(* IEC 61131-3 sources: plc-st-coding-agent/progress/v13_r8/upstream/datasets/public/tests, 2 files *)

(* ---- public-easy-04.reference.st ---- *)
(* Numeric millisecond variant of the jam-pump task. DebounceMs and CycleMs
   are in 1..3600000. No native TIME arithmetic is assumed. *)
FUNCTION_BLOCK FB
VAR_INPUT
    VISCOSITY_OK : BOOL;
    PASTE_E_STOP_NC : BOOL;
    DebounceMs : DINT;
    CycleMs : DINT;
END_VAR
VAR_OUTPUT
    VFD_RUN : BOOL;
    PUMP_MAINT_DUE : BOOL;
    PUMP_RUNTIME_ACC : LINT;
END_VAR
VAR
    validMs : DINT;
END_VAR

IF VISCOSITY_OK AND PASTE_E_STOP_NC THEN
    validMs := validMs + CycleMs;
    (* Durations beyond the largest permitted threshold are indistinguishable. *)
    IF validMs > 3600000 THEN
        validMs := 3600000;
    END_IF;
ELSE
    validMs := 0;
END_IF;
VFD_RUN := VISCOSITY_OK AND PASTE_E_STOP_NC AND validMs >= DebounceMs;
IF VFD_RUN THEN
    PUMP_RUNTIME_ACC := PUMP_RUNTIME_ACC + CycleMs;
END_IF;
PUMP_MAINT_DUE := PUMP_RUNTIME_ACC >= 1800000000;
END_FUNCTION_BLOCK

(* ---- public-medium-04.reference.st ---- *)
FUNCTION_BLOCK FB
VAR_INPUT
    TemperatureSensorInput : REAL;
    SetTemperature : REAL;
END_VAR
VAR_OUTPUT
    CurrentTemperature : REAL;
    SetTempDisplay : REAL;
    HeaterStatus : BOOL;
    OverheatProtection : BOOL;
    HeaterOutput : BOOL;
END_VAR
VAR
    onRun : INT;
    protectTimer : INT;
    fault : BOOL;
END_VAR

(* R6: 状态指示，当前温度与设定温度直通显示 *)
CurrentTemperature := TemperatureSensorInput;
SetTempDisplay := SetTemperature;

(* R7: 传感器故障判定：读数低于 0 或高于 100 视为故障 *)
fault := (TemperatureSensorInput < 0.0) OR (TemperatureSensorInput > 100.0);

IF OverheatProtection THEN
    (* R5: 过热保护期间强制关断加热；连续 3 拍（3s）冷却后解除 *)
    protectTimer := protectTimer + 1;
    IF protectTimer >= 3 THEN
        OverheatProtection := FALSE;
        protectTimer := 0;
        onRun := 0;
    ELSE
        HeaterOutput := FALSE;
    END_IF
END_IF

IF NOT OverheatProtection THEN
    (* R3/R4: 低于设定温度开加热，高于或等于设定温度关加热；
       传感器故障时禁止加热（R7 优先于 R3） *)
    IF fault THEN
        HeaterOutput := FALSE;
    ELSE
        HeaterOutput := TemperatureSensorInput < SetTemperature;
    END_IF

    (* R5: 连续加热计时，达到 5 拍（5s）即触发过热保护并立即关加热 *)
    IF HeaterOutput THEN
        onRun := onRun + 1;
        IF onRun >= 5 THEN
            OverheatProtection := TRUE;
            protectTimer := 0;
            onRun := 0;
            HeaterOutput := FALSE;
        END_IF
    ELSE
        onRun := 0;
    END_IF
END_IF

(* R6: 加热状态指示跟随实际加热输出 *)
HeaterStatus := HeaterOutput;
END_FUNCTION_BLOCK
